SUBAPPLICATION Sitzventile (* Subapplication Type *)
  (* Standard: 61499-2 *)
  (* Version 1.0, 2023-02-11, franz *)
  IMPORT logiBUS::io::DQ::logiBUS_DO::Invalid;
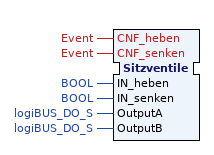
  EVENT_INPUT
    CNF_heben;
    CNF_senken;
  END_EVENT
  VAR_INPUT
    IN_heben : BOOL;
    IN_senken : BOOL;
    OutputA : logiBUS::io::DQ::logiBUS_DO_S := Invalid;
    OutputB : logiBUS::io::DQ::logiBUS_DO_S := Invalid;
  END_VAR
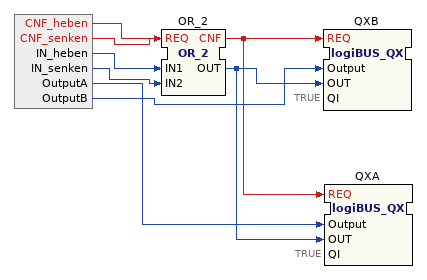
  FBS
    OR_2 : iec61131::bitwiseOperators::OR_2;
    QXB : logiBUS::io::DQ::logiBUS_QX(QI := TRUE);
    QXA : logiBUS::io::DQ::logiBUS_QX(QI := TRUE);
  END_FBS
  EVENT_CONNECTIONS
    OR_2.CNF TO QXB.REQ;
    OR_2.CNF TO QXA.REQ;
    CNF_heben TO OR_2.REQ;
    CNF_senken TO OR_2.REQ;
  END_CONNECTIONS
  DATA_CONNECTIONS
    OutputB TO QXB.Output;
    OutputA TO QXA.Output;
    OR_2.OUT TO QXB.OUT;
    OR_2.OUT TO QXA.OUT;
    IN_heben TO OR_2.IN1;
    IN_senken TO OR_2.IN2;
  END_CONNECTIONS
END_SUBAPPLICATION
